(* IEC 61131-3 sources: llm-plc-st-eval/data/processed_definitivo/claude-sonnet-4-6/B4/zero_shot, 3 files *)

(* ---- ejec_1.st ---- *)
FUNCTION_BLOCK FB_Giro
VAR_INPUT
    btnFwd  : BOOL; (* Botón marcha horaria *)
    btnRev  : BOOL; (* Botón marcha antihoraria *)
    btnParo : BOOL; (* Botón paro *)
END_VAR

VAR_OUTPUT
    fwd : BOOL; (* Salida giro horario *)
    rev : BOOL; (* Salida giro antihorario *)
END_VAR

VAR
    (* Estado interno: TRUE = en marcha, FALSE = parado *)
    xRunning : BOOL := FALSE;
END_VAR

(*
    Lógica de control:
    - btnParo detiene el motor (prioridad máxima).
    - btnFwd activa fwd solo si el motor está parado (rev = FALSE).
    - btnRev activa rev solo si el motor está parado (fwd = FALSE).
    - Nunca se permite cambio directo de sentido sin pasar por paro.
*)

(* ── 1. PARO: prioridad máxima ── *)
IF btnParo THEN
    fwd      := FALSE;
    rev      := FALSE;
    xRunning := FALSE;

(* ── 2. MARCHA HORARIA: solo si el motor está parado ── *)
ELSIF btnFwd AND NOT xRunning THEN
    fwd      := TRUE;
    rev      := FALSE;  (* Enclavamiento: rev siempre apagada *)
    xRunning := TRUE;

(* ── 3. MARCHA ANTIHORARIA: solo si el motor está parado ── *)
ELSIF btnRev AND NOT xRunning THEN
    rev      := TRUE;
    fwd      := FALSE;  (* Enclavamiento: fwd siempre apagada *)
    xRunning := TRUE;

(* ── 4. Sin pulsación relevante: mantener estado actual ── *)
END_IF;

(* ── 5. Enclavamiento de seguridad por hardware (doble seguro) ── *)
(* Garantiza que nunca ambas salidas estén activas, incluso ante  *)
(* corrupción de memoria o fallo lógico imprevisto.               *)
IF fwd AND rev THEN
    fwd      := FALSE;
    rev      := FALSE;
    xRunning := FALSE;
END_IF;

END_FUNCTION_BLOCK

(* ---- ejec_2.st ---- *)
FUNCTION_BLOCK FB_Giro
VAR_INPUT
    btnFwd  : BOOL; (* Botón marcha horaria *)
    btnRev  : BOOL; (* Botón marcha antihoraria *)
    btnParo : BOOL; (* Botón de paro *)
END_VAR

VAR_OUTPUT
    fwd : BOOL; (* Salida giro horario *)
    rev : BOOL; (* Salida giro antihorario *)
END_VAR

VAR
    (* Estado interno: TRUE = en marcha, FALSE = parado *)
    xRunning : BOOL := FALSE;
END_VAR

(*
    Lógica de control:
    - btnParo detiene el motor (prioridad alta).
    - btnFwd activa fwd solo si el motor está parado (xRunning = FALSE).
    - btnRev activa rev solo si el motor está parado (xRunning = FALSE).
    - Una vez en marcha, solo btnParo puede cambiar el estado.
    - fwd y rev nunca pueden estar activas simultáneamente.
*)

(* 1. Paro con prioridad máxima *)
IF btnParo THEN
    fwd      := FALSE;
    rev      := FALSE;
    xRunning := FALSE;

(* 2. Arranque en sentido horario: solo si el motor está parado *)
ELSIF btnFwd AND NOT xRunning THEN
    fwd      := TRUE;
    rev      := FALSE;  (* Interbloqueo: asegurar rev inactiva *)
    xRunning := TRUE;

(* 3. Arranque en sentido antihorario: solo si el motor está parado *)
ELSIF btnRev AND NOT xRunning THEN
    rev      := TRUE;
    fwd      := FALSE;  (* Interbloqueo: asegurar fwd inactiva *)
    xRunning := TRUE;

(* 4. Motor en marcha: mantener estado hasta recibir paro *)
(* No se hace nada; fwd/rev conservan su valor *)
END_IF;

(* 5. Interbloqueo de seguridad por hardware: nunca ambas activas *)
IF fwd AND rev THEN
    fwd      := FALSE;
    rev      := FALSE;
    xRunning := FALSE;
END_IF;

END_FUNCTION_BLOCK

(* ---- ejec_3.st ---- *)
FUNCTION_BLOCK FB_Giro
VAR_INPUT
    btnFwd  : BOOL; (* Botón marcha horaria *)
    btnRev  : BOOL; (* Botón marcha antihoraria *)
    btnParo : BOOL; (* Botón paro *)
END_VAR

VAR_OUTPUT
    fwd : BOOL; (* Salida giro horario *)
    rev : BOOL; (* Salida giro antihorario *)
END_VAR

VAR
    (* Estado interno: TRUE = en marcha, FALSE = parado *)
    xRunning : BOOL := FALSE;
END_VAR

(*
    Lógica de control:
    - btnParo detiene el motor (prioridad máxima).
    - btnFwd activa fwd solo si el motor está parado (rev = FALSE).
    - btnRev activa rev solo si el motor está parado (fwd = FALSE).
    - Nunca se permite activar fwd y rev simultáneamente.
    - Para invertir el giro es obligatorio pasar por paro.
*)

(* 1. Paro con prioridad máxima *)
IF btnParo THEN
    fwd      := FALSE;
    rev      := FALSE;
    xRunning := FALSE;

(* 2. Marcha horaria: solo si el motor está parado *)
ELSIF btnFwd AND NOT xRunning THEN
    fwd      := TRUE;
    rev      := FALSE;  (* Enclavamiento: garantiza rev = FALSE *)
    xRunning := TRUE;

(* 3. Marcha antihoraria: solo si el motor está parado *)
ELSIF btnRev AND NOT xRunning THEN
    rev      := TRUE;
    fwd      := FALSE;  (* Enclavamiento: garantiza fwd = FALSE *)
    xRunning := TRUE;

(* 4. Sin pulsación relevante: mantener estado actual *)
END_IF;
